(* CODESYS project controls.library
   DefaultNamespace: KOSTAL.AF2024.HMI.Controls
   DocFormat: reStructuredText
   Description: Provide functionalities of  HMI Controls
   Author: Frank Dümpelmann
   Title: KOSTAL.AF2024.HMI.Controls
   Version: 1.0.1.0
   Company: KOSTAL GmbH & Co.KG
   Placeholder: KOSTAL.AF2024.HMI.Controls

Project tree, tasks and I/O mapping:
  libraries: KOSTAL.AF2024.Core.Settings, 1.0.0.0 (KOSTAL GmbH & Co.KG); KOSTAL.AF2024.Core.System, 1.0.0.0 (KOSTAL GmbH & Co.KG)
  Button/
    interface I_T_Button: CopyTo, Pulse, Sign
    interface I_T_Button_CopyFrom: CopyFrom
    interface I_T_Button_Owner: clear, CopyFrom, CopyTo, Pulse, Sign
    function block T_Button [ST]: clear, CopyFrom, CopyTo, Pulse, Sign
  ButtonControlled/
    interface I_T_Button_controlled: clear_control, Text, Visible
    interface I_T_Button_controlled_Owner: clear_signals, Text, Visible
    interface I_T_Button_controlled_RO: Text, Visible
    function block T_Button_controlled [ST]: clear, clear_control, clear_signals, CopyFrom, Text, Visible
  Digital Input/
    function block FB_DigitalInput [ST]: clear, settings, Settings_RO, Signal
    interface I_DigitalInput: Settings_RO, Signal
    interface I_DigitalInput_Owner: clear, settings, Signal
  Digital Output/
    data type _ST_DoManual
    function block FB_DigitalOutput [ST]: _manualMode_Set, _manualModeControl, clear, clear_signal, FBmain, ManualMode_Reset, settings, settings_RO, Signal
    interface I_DigitalOutput: settings, Signal
    interface I_DigitalOutput_RO: settings_RO, Signal
  Project Information/
    function F_GetCompany [ST]
    function F_GetTitle [ST]
    function F_GetVersion [ST]
  Settings/
    interface I_T_settings: clear, CopyFrom, CopyTo, enable, name
    interface I_T_settings_CopyFrom: CopyFrom
    interface I_T_settings_RO: enable, name
    function block T_settings [ST]: clear, CopyFrom, CopyTo, enable, name
  Text/
    interface I_T_text: CopyTo, text
    interface I_T_text_CopyFrom: CopyFrom
    function block T_text [ST]: clear, CopyFrom, CopyTo, text
  Version/
    global variables Global_Version
*)

// Digital Output/_ST_DoManual

TYPE _ST_DoManual :
STRUCT
	ManualMode 	: BOOL;
	ManualInterlock 	: BOOL;
	AutomaticRelease 	: BOOL;
	
	RequestManualOn		: BOOL;
	RequestManualOff	: BOOL;
	
	Sign				: BOOL;
	ResetCounter		: BYTE := 1;
	
END_STRUCT
END_TYPE

// Version/Global_Version
{attribute 'TcGenerated'}
{attribute 'no-analysis'}
{attribute 'linkalways'}
// This function has been automatically generated from the project information.
VAR_GLOBAL CONSTANT
	{attribute 'const_non_replaced'}
	stLibVersion_KOSTAL_AF2024_HMI_Controls : ST_LibVersion := (iMajor := 1, iMinor := 0, iBuild := 1, iRevision := 0, nFlags := 0, sVersion := '1.0.1.0');
END_VAR

// Button/I_T_Button
INTERFACE I_T_Button EXTENDS KOSTAL_AF2024_Core_System.I_Interface

METHOD PUBLIC CopyTo
VAR_INPUT
	IN	: I_T_Button_CopyFrom;
END_VAR
END_METHOD

(*
Description
===========
| TRUE for one cycle when the button is pressed
*)
PROPERTY PUBLIC Pulse : BOOL
GET
END_GET
END_PROPERTY

(*
Description
===========
| TRUE while the button is pressed
*)
PROPERTY PUBLIC Sign : BOOL
GET
END_GET
END_PROPERTY

END_INTERFACE

// Button/I_T_Button_CopyFrom
INTERFACE I_T_Button_CopyFrom EXTENDS KOSTAL_AF2024_Core_System.I_Interface

METHOD PUBLIC CopyFrom
VAR_INPUT
	IN	: I_T_Button;
END_VAR
END_METHOD

END_INTERFACE

// Button/I_T_Button_Owner
INTERFACE I_T_Button_Owner EXTENDS KOSTAL_AF2024_Core_System.I_Interface

(*
Description
===========
| Reset signals
*)
METHOD PUBLIC clear
END_METHOD

METHOD PUBLIC CopyFrom
VAR_INPUT
	IN	: I_T_Button;
END_VAR
END_METHOD

METHOD PUBLIC CopyTo
VAR_INPUT
	IN	: I_T_Button_CopyFrom;
END_VAR
END_METHOD

(*
Description
===========
| TRUE for one cycle when the button is pressed
*)
PROPERTY PUBLIC Pulse : BOOL
GET
END_GET
SET
END_SET
END_PROPERTY

(*
Description
===========
| TRUE while the button is pressed
*)
PROPERTY PUBLIC Sign : BOOL
GET
END_GET
SET
END_SET
END_PROPERTY

END_INTERFACE

// Button/T_Button
(*

:Author: Frank Dümpelmann <f.duempelmann@kostal.com>, Martin Hundt <m.hundt@kostal.com>
:Date: 2018-11-20

Function
========
Data structure representing the signals of an HMI button 

Usage notes
===============
| To be used in HMI application , such as TP57AT
*)
FUNCTION_BLOCK PUBLIC T_Button IMPLEMENTS I_T_Button, I_T_Button_Owner, I_T_Button_CopyFrom

VAR
	_Sign		: BOOL;	//BOOL
	_Pulse	: BOOL;	//BOOL
END_VAR

(*
Description
===========
| Reset signals
*)
METHOD PUBLIC clear

_Sign	:= FALSE;
_Pulse:= FALSE;
END_METHOD

METHOD PUBLIC CopyFrom
VAR_INPUT
	IN	: I_T_Button;
END_VAR

IF IN = 0 THEN RETURN;	END_IF

_Pulse	:= IN.Pulse;
_Sign		:= IN.Sign;
END_METHOD

METHOD PUBLIC CopyTo
VAR_INPUT
	IN	: I_T_Button_CopyFrom;
END_VAR

IF IN = 0 THEN RETURN;	END_IF

IN.CopyFrom(THIS^);
END_METHOD

(*
Description
===========
| TRUE for one cycle when the button is pressed
*)
PROPERTY PUBLIC Pulse : BOOL
GET

Pulse:= _Pulse;
END_GET
SET

_Pulse:= Pulse;
END_SET
END_PROPERTY

(*
Description
===========
| TRUE while the button is pressed
*)
PROPERTY PUBLIC Sign : BOOL
GET

Sign:= _Sign;
END_GET
SET

_Sign:= Sign;
END_SET
END_PROPERTY

END_FUNCTION_BLOCK

// ButtonControlled/I_T_Button_controlled
INTERFACE I_T_Button_controlled EXTENDS I_T_Button_controlled_RO

METHOD PUBLIC clear_control
END_METHOD

PROPERTY PUBLIC Text : WSTRING(40)
SET
END_SET
END_PROPERTY

PROPERTY PUBLIC Visible : BOOL
SET
END_SET
END_PROPERTY

END_INTERFACE

// ButtonControlled/I_T_Button_controlled_RO
INTERFACE I_T_Button_controlled_RO EXTENDS I_T_Button

PROPERTY PUBLIC Text : WSTRING(40)
GET
END_GET
END_PROPERTY

PROPERTY PUBLIC Visible : BOOL
GET
END_GET
END_PROPERTY

END_INTERFACE

// ButtonControlled/I_T_Button_controlled_Owner
INTERFACE I_T_Button_controlled_Owner EXTENDS I_T_Button_Owner

METHOD PUBLIC clear_signals
END_METHOD

PROPERTY PUBLIC Text : WSTRING(40)
GET
END_GET
SET
END_SET
END_PROPERTY

PROPERTY PUBLIC Visible : BOOL
GET
END_GET
SET
END_SET
END_PROPERTY

END_INTERFACE

// ButtonControlled/T_Button_controlled
(*

:Author: Frank Dümpelmann <f.duempelmann@kostal.com>, Martin Hundt <m.hundt@kostal.com>
:Date: 2018-11-20

Function
========
| Data structure representing an HMI button 

Usage notes
===============
| To be used in HMI application , such as TP57AT

Methods and Properties
======================
| clear: clear all content and signals
| clear_signals: clear signals (button pushed) only
| Text and visibility of the button
| See documentation of FB_Button for inherited methods and properties

*)
FUNCTION_BLOCK PUBLIC T_Button_controlled EXTENDS T_Button IMPLEMENTS I_T_Button_controlled_RO, I_T_Button_controlled_Owner, I_T_Button_controlled

VAR
	_Visible	: BOOL;
	_Text			: WSTRING;
END_VAR

METHOD PUBLIC clear

SUPER^.clear();

_Visible:= FALSE;
_Text		:= "";
END_METHOD

METHOD PUBLIC clear_control

_Visible:= FALSE;
_Text		:= "";
END_METHOD

METHOD PUBLIC clear_signals

SUPER^.clear();
END_METHOD

METHOD PUBLIC CopyFrom
VAR_INPUT
	IN	: I_T_Button;
END_VAR

VAR
	_obj	: I_T_Button_controlled_RO:= 0;
END_VAR

IF IN = 0 THEN RETURN;	END_IF

IF NOT __QUERYINTERFACE(IN, _obj) THEN RETURN; END_IF
IF _obj = 0 THEN RETURN;	END_IF

_Visible	:= _obj.Visible;
_Text			:= _obj.Text;

SUPER^.CopyFrom(IN);
END_METHOD

PROPERTY PUBLIC Text : WSTRING(40)
GET

Text:= _Text;
END_GET
SET

_Text:= Text;
END_SET
END_PROPERTY

PROPERTY PUBLIC Visible : BOOL
GET

Visible:= _Visible;
END_GET
SET

_Visible:= Visible;
END_SET
END_PROPERTY

END_FUNCTION_BLOCK

// Digital Input/FB_DigitalInput
(*

:Author: Frank Dümpelmann <f.duempelmann@kostal.com>, Martin Hundt <m.hundt@kostal.com>
:Date: 2018-11-20

Function
========
Data type representing a digital input (sensor etc.)

Methods and Properties
======================
| Signal: Signal of the sensor
| settings: see T_settings
| clear: clear settings

*)
FUNCTION_BLOCK PUBLIC FB_DigitalInput IMPLEMENTS I_DigitalInput, I_DigitalInput_Owner

VAR
	{attribute 'DigitalInput_2024_V1'}
	_settings		: T_settings;	//FB_sensor_settings
	input	 AT %I*	: BOOL;		//BOOL
END_VAR

METHOD PUBLIC clear
VAR_INPUT
END_VAR

_settings.clear();
END_METHOD

PROPERTY PUBLIC settings : I_T_settings
GET

settings := _settings;
END_GET
END_PROPERTY

PROPERTY PUBLIC Settings_RO : I_T_settings_RO
GET

Settings_RO:= _settings;
END_GET
END_PROPERTY

PROPERTY PUBLIC Signal : BOOL
GET

Signal:= input;
END_GET
END_PROPERTY

END_FUNCTION_BLOCK

// Settings/T_settings
(*

:Author: Frank Dümpelmann <f.duempelmann@kostal.com>, Martin Hundt <m.hundt@kostal.com>
:Date: 2018-11-20

Function
========
Data type representing a sensor's settings

Methods and Properties
======================
| Name of the sensor, enable/disable, clear all
*)
FUNCTION_BLOCK PUBLIC T_settings IMPLEMENTS I_T_settings_RO, I_T_settings_CopyFrom, I_T_settings

VAR
	_enable	: BOOL;		//BOOL
	_name		: KOSTAL_AF2024_Core_Settings.T_MaxString;	//STRING
END_VAR

METHOD PUBLIC clear
VAR_INPUT
END_VAR


_enable	:= FALSE;
_name		:= "";
END_METHOD

METHOD PUBLIC CopyFrom
VAR_INPUT
	IN	: I_T_settings_RO;
END_VAR

IF IN = 0 THEN RETURN;	END_IF

_enable	:= IN.enable;
_name		:= IN.name;
END_METHOD

METHOD PUBLIC CopyTo
VAR_INPUT
	IN	: I_T_settings_CopyFrom;
END_VAR

IF IN = 0 THEN RETURN;	END_IF

IN.CopyFrom(THIS^);
END_METHOD

PROPERTY PUBLIC enable : BOOL
GET

enable:= _enable;
END_GET
SET

_enable:= enable;
END_SET
END_PROPERTY

PROPERTY PUBLIC name : KOSTAL_AF2024_Core_Settings.T_MaxString
GET

name:= _name;
END_GET
SET

_name:= name;
END_SET
END_PROPERTY

END_FUNCTION_BLOCK

// Settings/I_T_settings_RO
INTERFACE I_T_settings_RO EXTENDS KOSTAL_AF2024_Core_System.I_Interface

PROPERTY PUBLIC enable : BOOL
GET
END_GET
END_PROPERTY

PROPERTY PUBLIC name : KOSTAL_AF2024_Core_Settings.T_MaxString
GET
END_GET
END_PROPERTY

END_INTERFACE

// Settings/I_T_settings_CopyFrom
INTERFACE I_T_settings_CopyFrom EXTENDS KOSTAL_AF2024_Core_System.I_Interface

METHOD PUBLIC CopyFrom
VAR_INPUT
	IN	: I_T_settings_RO;
END_VAR
END_METHOD

END_INTERFACE

// Settings/I_T_settings
INTERFACE I_T_settings EXTENDS KOSTAL_AF2024_Core_System.I_Interface

METHOD PUBLIC clear
VAR_INPUT
END_VAR
END_METHOD

METHOD PUBLIC CopyFrom
VAR_INPUT
	IN	: I_T_settings_RO;
END_VAR
END_METHOD

METHOD PUBLIC CopyTo
VAR_INPUT
	IN	: I_T_settings_CopyFrom;
END_VAR
END_METHOD

PROPERTY PUBLIC enable : BOOL
GET
END_GET
SET
END_SET
END_PROPERTY

PROPERTY PUBLIC name : KOSTAL_AF2024_Core_Settings.T_MaxString
GET
END_GET
SET
END_SET
END_PROPERTY

END_INTERFACE

// Digital Input/I_DigitalInput
INTERFACE I_DigitalInput EXTENDS KOSTAL_AF2024_Core_System.I_Interface

PROPERTY PUBLIC Settings_RO : I_T_settings_RO
GET
END_GET
END_PROPERTY

PROPERTY PUBLIC Signal : BOOL
GET
END_GET
END_PROPERTY

END_INTERFACE

// Digital Input/I_DigitalInput_Owner
INTERFACE I_DigitalInput_Owner EXTENDS KOSTAL_AF2024_Core_System.I_Interface

METHOD PUBLIC clear
VAR_INPUT
END_VAR
END_METHOD

PROPERTY PUBLIC settings : I_T_settings
GET
END_GET
END_PROPERTY

PROPERTY PUBLIC Signal : BOOL
GET
END_GET
END_PROPERTY

END_INTERFACE

// Digital Output/FB_DigitalOutput
(*

:Author: Martin Hundt <m.hundt@kostal.com>
:Date: 2023-07-20

Function
========
| Function Block representing a digital output
| Interface for manual control from HMI


Methods and Properties
======================
| Signal: Signal of the sensor
| settings: see T_settings
| clear: clear all
| clear_sign: clear signal only

*)
FUNCTION_BLOCK PUBLIC FB_DigitalOutput IMPLEMENTS I_DigitalOutput, I_DigitalOutput_RO

VAR
	_settings			: T_settings;	
	_sign				: BOOL;		//BOOL
	output		AT %Q* 	: BOOL;		//BOOL
	
	{attribute 'DigitalOutput_2024_V1'}
	_manual		: _ST_DoManual;
END_VAR

(*
Description
===========
| (De)activate manual valve mode
| Parameters:
| 	state : bool : TRUE = activate, FALSE = deactivate
*)
METHOD PROTECTED _manualMode_Set
VAR_INPUT
	state : bool;
END_VAR
IF state THEN
	_manual.ManualMode := TRUE;
ELSE
	_manual.ManualMode 	:= FALSE;
END_IF
END_METHOD

METHOD PROTECTED _manualModeControl
VAR_INPUT
END_VAR
_manual.AutomaticRelease := (output = _sign);

IF _manual.RequestManualOn AND NOT _manual.ManualInterlock AND NOT _manual.ManualMode THEN
	_manualMode_Set(TRUE);
ELSIF _manual.RequestManualOff AND _manual.AutomaticRelease AND _manual.ManualMode THEN
	_manualMode_Set(FALSE);
END_IF

IF _manual.ManualMode AND NOT _manual.ManualInterlock THEN
	output := _manual.Sign;
ELSE
	output := _sign;
END_IF
END_METHOD

METHOD PUBLIC clear
VAR_INPUT
END_VAR
clear_signal();
_settings.clear();
END_METHOD

METHOD PUBLIC clear_signal
VAR_INPUT
END_VAR

_sign:= FALSE;
END_METHOD

METHOD PUBLIC FBmain
VAR_INPUT
END_VAR
_manualModeControl();
END_METHOD

METHOD PUBLIC ManualMode_Reset : BOOL
VAR_INPUT
END_VAR

_manualMode_Set(FALSE);
_manual.Sign := FALSE;
_manual.ResetCounter := LIMIT(1, _manual.ResetCounter + 1, 254);

_sign := false;
output := _sign;
END_METHOD

PROPERTY PUBLIC settings : I_T_settings
GET

settings := _settings;
END_GET
END_PROPERTY

PROPERTY PUBLIC settings_RO : I_T_settings_RO
GET

settings_RO := _settings;
END_GET
END_PROPERTY

PROPERTY PUBLIC Signal : BOOL
GET

Signal:= _sign;
END_GET
SET

_sign:= Signal;
END_SET
END_PROPERTY

END_FUNCTION_BLOCK

// Digital Output/I_DigitalOutput
INTERFACE I_DigitalOutput EXTENDS __SYSTEM.IQueryInterface

PROPERTY PUBLIC settings : I_T_settings
GET
END_GET
END_PROPERTY

PROPERTY PUBLIC Signal : BOOL
GET
END_GET
SET
END_SET
END_PROPERTY

END_INTERFACE

// Digital Output/I_DigitalOutput_RO
INTERFACE I_DigitalOutput_RO EXTENDS __SYSTEM.IQueryInterface

PROPERTY PUBLIC settings_RO : I_T_settings_RO
GET
END_GET
END_PROPERTY

PROPERTY PUBLIC Signal : BOOL
GET
END_GET
END_PROPERTY

END_INTERFACE

// Project Information/F_GetCompany
// This function has been automatically generated from the project information.
{attribute 'signature_flag' := '1073741824'}
{attribute 'TcGenerated'}
{attribute 'no-analysis'}
FUNCTION F_GetCompany : WSTRING
VAR_INPUT
	
END_VAR

F_GetCompany := "KOSTAL GmbH & Co.KG";

END_FUNCTION

// Project Information/F_GetTitle
// This function has been automatically generated from the project information.
{attribute 'signature_flag' := '1073741824'}
{attribute 'TcGenerated'}
{attribute 'no-analysis'}
FUNCTION F_GetTitle : WSTRING
VAR_INPUT
	
END_VAR

F_GetTitle := "KOSTAL.AF2024.HMI.Controls";

END_FUNCTION

// Project Information/F_GetVersion
// This function has been automatically generated from the project information.
{attribute 'signature_flag' := '1073741824'}
{attribute 'TcGenerated'}
{attribute 'no-analysis'}
FUNCTION F_GetVersion : ST_LibVersion
VAR_INPUT
	
END_VAR

F_GetVersion.iMajor := 1;
F_GetVersion.iMinor := 0;
F_GetVersion.iBuild := 1;
F_GetVersion.iRevision := 0;
F_GetVersion.sVersion := '1.0.1.0';
F_GetVersion.nFlags := 0;

END_FUNCTION

// Text/I_T_text
INTERFACE I_T_text EXTENDS __SYSTEM.IQueryInterface

METHOD PUBLIC CopyTo
VAR_INPUT
	IN	: I_T_text_CopyFrom;
END_VAR
END_METHOD

PROPERTY PUBLIC text : KOSTAL_AF2024_Core_Settings.T_MaxString
GET
END_GET
END_PROPERTY

END_INTERFACE

// Text/I_T_text_CopyFrom
INTERFACE I_T_text_CopyFrom

METHOD PUBLIC CopyFrom
VAR_INPUT
	IN	: I_T_text;
END_VAR
END_METHOD

END_INTERFACE

// Text/T_text
(*
| base class for text object
*)
FUNCTION_BLOCK PUBLIC T_text IMPLEMENTS I_T_text, I_T_text_CopyFrom

VAR
	_text	: KOSTAL_AF2024_Core_Settings.T_MaxString;
END_VAR

METHOD PUBLIC clear
VAR_INPUT
END_VAR

_text:= "";
END_METHOD

METHOD PUBLIC CopyFrom
VAR_INPUT
	IN	: I_T_text;
END_VAR

IF IN = 0 THEN RETURN;	END_IF

_text:= IN.text;
END_METHOD

METHOD PUBLIC CopyTo
VAR_INPUT
	IN	: I_T_text_CopyFrom;
END_VAR

IF IN = 0 THEN RETURN;	END_IF

IN.CopyFrom(THIS^);
END_METHOD

PROPERTY PUBLIC text : KOSTAL_AF2024_Core_Settings.T_MaxString
GET

text:= _text;
END_GET
SET

_text:= text;
END_SET
END_PROPERTY

END_FUNCTION_BLOCK
